{attribute 'call_after_init'}
FUNCTION_BLOCK FB_MyTimingSample
VAR
    nTimestampFB_init   : Tc2_EtherCAT.T_DCTIME64;
    nTimestampFB_reinit : Tc2_EtherCAT.T_DCTIME64;
    nTimestampMyInit    : Tc2_EtherCAT.T_DCTIME64;
END_VAR

METHOD FB_init : BOOL
VAR_INPUT
    bInitRetains : BOOL;
    bInCopyCode  : BOOL;
END_VAR
nTimestampFB_init := Tc2_EtherCAT.F_GetActualDcTime64();
FB_init := TRUE;
END_METHOD

METHOD FB_reinit : BOOL
VAR_INPUT
END_VAR
nTimestampFB_reinit := Tc2_EtherCAT.F_GetActualDcTime64();
FB_reinit := TRUE;
END_METHOD

{attribute 'call_after_init'}
METHOD MyInit : BOOL
nTimestampMyInit := Tc2_EtherCAT.F_GetActualDcTime64();
MyInit := TRUE;
END_METHOD

END_FUNCTION_BLOCK

(* stored: Version 1.1.0.1, ProductVersion 3.1.4024.16
   POU FB_MyTimingSample: Id {9cbe05af-01a4-4d3c-b0e3-9046fa23a359}, SpecialFunc None
   Method FB_init: Id {2a55bf74-edf4-42d1-b74c-77ebbb937d90}
   Method FB_reinit: Id {57537796-dc9e-4b87-bf7b-aa51f9c09a10}
   Method MyInit: Id {20688810-ad08-442d-b284-aeca832cb7ed} *)
